Fanuc KAREL source: ko00034.KL

-- PROVISIONAL review KL for V1013-1; original PC SHA256 bf4ae88c28de4419d830b5fc1aa02298c1667c9b52ec2288a39d350ebd2ab773
-- Incomplete behavior may be omitted. Consult companion uncertainty JSON. Do not deploy.
PROGRAM KO00034
%NOLOCKGROUP
BEGIN
  -- UNRESOLVED_PC offsets 5-12; opcodes 9D,23
  -- UNRESOLVED_PC offsets 17-66; opcodes 27,27,49,7E,AD,22,1C,22,31,7E,4A
  -- UNRESOLVED_PC offsets 71-75; opcodes 7F
END KO00034
